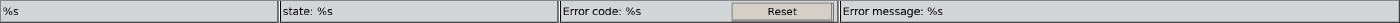
VISUALIZATION vis_Device_Error  // 1500x25
VAR_IN_OUT
	fb_comm_dev: fb_common_device;
END_VAR
    Rectangle (900,0 600x25), "Error message: %s", text variable: fb_comm_dev.common_events.device_error.error_string, colour toggle: fb_comm_dev.common_events.device_error.error_code<>''
        OnMouseUp: execute { GVL.Errors:=(0); }
    Rectangle (600,0 298x25), "Error code: %s", text variable: fb_comm_dev.common_events.device_error.error_code, colour toggle: fb_comm_dev.common_events.device_error.error_code<>''
        OnMouseUp: execute { GVL.Errors:=(0); }
    Button (784,3 109x20), "Reset"
        toggle fb_comm_dev.common_actions.reset
    Rectangle (0,0 298x25), "%s", tooltip "Device Name", text variable: fb_comm_dev.Name, colour toggle: fb_comm_dev.common_events.device_error.error_code<>''
        OnMouseUp: execute { GVL.Errors:=(0); }
    Rectangle (300,0 298x25), "state: %s", tooltip "Device State", text variable: fb_comm_dev.device_status, colour toggle: fb_comm_dev.common_events.device_error.error_code<>''
        OnMouseUp: execute { GVL.Errors:=(0); }
END_VISUALIZATION

(* stored: Version 1.1.0.1, ProductVersion 3.1.4024.12
   Visu vis_Device_Error: Id {90067ef6-653f-4908-b7f4-dfc056d70718} *)
